(* IEC 61131-3 sources: plcassist-cli/packages/volt-lsp-iec/test-corpus/twincat-project14/References/Tc3_Module, 38 files *)

(* ---- Global_Version.gvl ---- *)
VAR_GLOBAL
	stLibVersion_Tc3_Module : ST_LibVersion;
END_VAR

(* ---- GVL.gvl ---- *)
VAR_GLOBAL
	S_OK : HRESULT;
	S_FALSE : HRESULT;
	S_PENDING : HRESULT;
	S_WATCHDOG_TIMEOUT : HRESULT;
	E_FAIL : HRESULT;
	ERR_INVALID_PARAM : HRESULT;
	OTCID_CreateNewId : OTCID;
	OTCID_FirstFreeId : OTCID;
	OTCID_LastFreeId : OTCID;
	NULL : PVOID;
END_VAR

(* ---- ExCpHndFunc.fun ---- *)
FUNCTION ExCpHndFunc : UDINT
VAR_INPUT
	pUsr : PVOID;
	pExcpHndPara : PVOID;
END_VAR
END_FUNCTION

(* ---- F_CPUCounter.fun ---- *)
FUNCTION F_CPUCounter : BOOL
VAR_INPUT
	counter : ULINT;
END_VAR
END_FUNCTION

(* ---- F_TcLicSrv_TakeLicense.fun ---- *)
FUNCTION F_TcLicSrv_TakeLicense : HRESULT
VAR_INPUT
	refLicenseId : REFERENCE TO GUID;
END_VAR
END_FUNCTION

(* ---- FAILED.fun ---- *)
FUNCTION FAILED : BOOL
VAR_INPUT
	hr : HRESULT;
END_VAR
END_FUNCTION

(* ---- FW_GetAppState.fun ---- *)
FUNCTION FW_GetAppState : UDINT
END_FUNCTION

(* ---- FW_MemCmp.fun ---- *)
FUNCTION FW_MemCmp : DINT
VAR_INPUT
	pBuf1 : PVOID;
	pBuf2 : PVOID;
	cbLen : UDINT;
END_VAR
END_FUNCTION

(* ---- FW_MemCpy.fun ---- *)
FUNCTION FW_MemCpy : UDINT
VAR_INPUT
	pDest : PVOID;
	pSrc : PVOID;
	cbLen : UDINT;
END_VAR
END_FUNCTION

(* ---- FW_MemSet.fun ---- *)
FUNCTION FW_MemSet : UDINT
VAR_INPUT
	pDest : PVOID;
	nFillByte : USINT;
	cbLen : UDINT;
END_VAR
END_FUNCTION

(* ---- FW_ObjMgr_CreateAndInitInstance.fun ---- *)
FUNCTION FW_ObjMgr_CreateAndInitInstance : HRESULT
VAR_INPUT
	clsId : CLSID;
	iid : IID;
	pipUnk : POINTER TO ITcUnknown;
	objId : UDINT;
	parentId : UDINT;
	name : REFERENCE TO STRING;
	state : UDINT;
	pInitData : POINTER TO TComInitDataHdr;
END_VAR
END_FUNCTION

(* ---- FW_ObjMgr_CreateInstance.fun ---- *)
FUNCTION FW_ObjMgr_CreateInstance : HRESULT
VAR_INPUT
	clsId : CLSID;
	iid : IID;
	pipUnk : POINTER TO ITcUnknown;
END_VAR
END_FUNCTION

(* ---- FW_ObjMgr_DeleteInstance.fun ---- *)
FUNCTION FW_ObjMgr_DeleteInstance : HRESULT
VAR_INPUT
	pipUnk : POINTER TO ITcUnknown;
END_VAR
END_FUNCTION

(* ---- FW_ObjMgr_DeregisterObject.fun ---- *)
FUNCTION FW_ObjMgr_DeregisterObject : HRESULT
VAR_INPUT
	oidApp : OTCID;
	oidObj : OTCID;
	bInCopyCode : BOOL;
END_VAR
END_FUNCTION

(* ---- FW_ObjMgr_GetObjectInstance.fun ---- *)
FUNCTION FW_ObjMgr_GetObjectInstance : HRESULT
VAR_INPUT
	oid : OTCID;
	iid : IID;
	pipUnk : POINTER TO ITcUnknown;
END_VAR
END_FUNCTION

(* ---- FW_ObjMgr_GetObjectServer.fun ---- *)
FUNCTION FW_ObjMgr_GetObjectServer : HRESULT
VAR_INPUT
	oidApp : OTCID;
	pipSrv : POINTER TO ITComObjectServer;
END_VAR
END_FUNCTION

(* ---- FW_ObjMgr_RegisterObject.fun ---- *)
FUNCTION FW_ObjMgr_RegisterObject : HRESULT
VAR_INPUT
	oidApp : OTCID;
	oidObj : OTCID;
	bInCopyCode : BOOL;
	ipUnk : ITcUnknown;
END_VAR
END_FUNCTION

(* ---- FW_SafeRelease.fun ---- *)
FUNCTION FW_SafeRelease : HRESULT
VAR_INPUT
	pipUnk : POINTER TO ITcUnknown;
END_VAR
END_FUNCTION

(* ---- Fw_Trace.fun ---- *)
FUNCTION Fw_Trace : DINT
VAR_INPUT
	val : DINT;
	text : STRING(255);
END_VAR
END_FUNCTION

(* ---- GuidsEqual.fun ---- *)
FUNCTION GuidsEqual : BOOL
VAR_INPUT
	pGuidA : POINTER TO GUID;
	pGuidB : POINTER TO GUID;
END_VAR
END_FUNCTION

(* ---- ITCUNKNOWN_TO_PVOID.fun ---- *)
FUNCTION ITCUNKNOWN_TO_PVOID : PVOID
VAR_INPUT
	itcUnknown : ITcUnknown;
END_VAR
END_FUNCTION

(* ---- MEMCMP.fun ---- *)
FUNCTION MEMCMP : DINT
VAR_INPUT
	pBuf1 : PVOID;
	pBuf2 : PVOID;
	n : UDINT;
END_VAR
END_FUNCTION

(* ---- MEMCPY.fun ---- *)
FUNCTION MEMCPY : UDINT
VAR_INPUT
	destAddr : PVOID;
	srcAddr : PVOID;
	n : UDINT;
END_VAR
END_FUNCTION

(* ---- MEMSET.fun ---- *)
FUNCTION MEMSET : UDINT
VAR_INPUT
	destAddr : PVOID;
	fillByte : USINT;
	n : UDINT;
END_VAR
END_FUNCTION

(* ---- POINTERTOINTERFACE_TO_PVOID.fun ---- *)
FUNCTION POINTERTOINTERFACE_TO_PVOID : PVOID
VAR_INPUT
	pTmp : POINTER TO PVOID;
END_VAR
END_FUNCTION

(* ---- PTComInitDataElmHdrDATA.fun ---- *)
FUNCTION PTComInitDataElmHdrDATA : POINTER TO TComInitDataElmHdr
VAR_INPUT
	pTComInitDataElmHdr : POINTER TO TComInitDataElmHdr;
END_VAR
END_FUNCTION

(* ---- PTComInitDataElmHdrNEXTHDR.fun ---- *)
FUNCTION PTComInitDataElmHdrNEXTHDR : POINTER TO TComInitDataElmHdr
VAR_INPUT
	pTComInitDataElmHdr : POINTER TO TComInitDataElmHdr;
END_VAR
END_FUNCTION

(* ---- PTComInitDataElmHdrSIZEOF.fun ---- *)
FUNCTION PTComInitDataElmHdrSIZEOF : DINT
VAR_INPUT
	pTComInitDataElmHdr : POINTER TO TComInitDataElmHdr;
END_VAR
END_FUNCTION

(* ---- PVOID_TO_ITCUNKNOWN.fun ---- *)
FUNCTION PVOID_TO_ITCUNKNOWN : ITcUnknown
VAR_INPUT
	pVoid : PVOID;
END_VAR
END_FUNCTION

(* ---- PVOID_TO_POINTERTOINTERFACE.fun ---- *)
FUNCTION PVOID_TO_POINTERTOINTERFACE : POINTER TO ITcUnknown
VAR_INPUT
	pVoid : PVOID;
END_VAR
END_FUNCTION

(* ---- SizeOfCString.fun ---- *)
FUNCTION SizeOfCString : UDINT
VAR_INPUT
	myCString : POINTER TO STRING;
END_VAR
END_FUNCTION

(* ---- SUCCEEDED.fun ---- *)
FUNCTION SUCCEEDED : BOOL
VAR_INPUT
	hr : HRESULT;
END_VAR
END_FUNCTION

(* ---- TaskFnc.fun ---- *)
FUNCTION TaskFnc : UDINT
VAR_INPUT
	pUsr : PVOID;
END_VAR
END_FUNCTION

(* ---- IecTaskModule.fb ---- *)
FUNCTION_BLOCK IecTaskModule
END_FUNCTION_BLOCK

(* ---- IecTaskModulePost.fb ---- *)
FUNCTION_BLOCK IecTaskModulePost
END_FUNCTION_BLOCK

(* ---- TcBaseModule.fb ---- *)
FUNCTION_BLOCK TcBaseModule
END_FUNCTION_BLOCK

(* ---- TcBaseModuleRegistered.fb ---- *)
FUNCTION_BLOCK TcBaseModuleRegistered
END_FUNCTION_BLOCK

(* ---- TcBaseModuleRegistered2.fb ---- *)
FUNCTION_BLOCK TcBaseModuleRegistered2
VAR_OUTPUT
	objID : OTCID;
END_VAR
END_FUNCTION_BLOCK
